# EPICS substitutions: db/Beckhoff_7XXX/ecmcEP7211-0034_OPT_info2Inputs.substitutions
file "ecmcEP7211-0034_INFO2_INPUTS.template"
{
  pattern {CH_ID}
          {01   }
}
